FUNCTION_BLOCK "naut_Slow"
{ S7_Optimized_Access := 'TRUE' }
VERSION : 0.1
   VAR
      i : INT;
   END_VAR
   VAR_TEMP
      naut_for_v1 : INT;
   END_VAR

BEGIN
	"naut_Scan_slow".tags.Status.%X3 := "naut_Scan_slow".tags.Level > 10.0;
	"naut_Scan_slow".assigned.Status.%X3 := TRUE;
	IF "naut_Scan_slow".tags.Stop THEN
		"naut_Scan_slow".tags.Status.%X0 := TRUE;
		"naut_Scan_slow".assigned.Status.%X0 := TRUE;
	END_IF;
	IF "naut_Scan_slow".tags.Start THEN
		"naut_Scan_slow".tags.Status := 16#0;
		"naut_Scan_slow".assigned.Status := WORD#16#FFFF;
	END_IF;
	FOR #naut_for_v1 := 1 TO 3 DO
		#i := #naut_for_v1;
		"naut_Scan_slow".tags.Status.%X7 := NOT "naut_Scan_slow".tags.Status.%X7;
		"naut_Scan_slow".assigned.Status.%X7 := TRUE;
	END_FOR;
	#i := 4;
END_FUNCTION_BLOCK
